Staubli VAL3: main.pgx

public program main()
begin
  //start
  call iolink()

  //main loop
  do
    call safePointCheck()


    call safeZoneCheck()


    delay(0)
  until false
end
